(* PLC project g_busbar_interlock_clean, Anonymous Benchmark Suite 1.0 *)
(* stored: creationDateTime 2026-07-09T00:00:00 *)

PROGRAM g_busbar_interlock_clean
  VAR_INPUT
    feeder_a_cmd : BOOL;
    feeder_b_cmd : BOOL;
    maint : BOOL;
  END_VAR
  VAR_OUTPUT
    feeder_a : BOOL;
    feeder_b : BOOL;
  END_VAR

(* LD diagram, written out as Structured Text *)
feeder_a := NOT feeder_b_cmd AND feeder_a_cmd;
feeder_b := feeder_b_cmd;
END_PROGRAM

CONFIGURATION Config0
  RESOURCE Res0 ON PLC
    TASK tcyclic(INTERVAL := T#10ms, PRIORITY := 0);
    PROGRAM inst0 WITH tcyclic : g_busbar_interlock_clean;
  END_RESOURCE
END_CONFIGURATION
